    "FRK_Line".Data.BuiltRevision := "FRK_Line".Data.Status.Revision;
    #FRK_DocApply_D011 := TRUE;
END_FUNCTION
FUNCTION "FRK_DocCapture_D012" : Bool
{ S7_Optimized_Access := 'TRUE' }
VERSION : 0.1
VAR_IN_OUT
    Length : DInt;
END_VAR
VAR_TEMP
    Index : Int;
    Stored : Int;
    Position : DInt;
    NativeResult : Int;
    Ok : Bool;
END_VAR
BEGIN
    #FRK_DocCapture_D012 := FALSE;
    "FRK_PersistImages".D012.SchemaVersion := 1; "FRK_PersistImages".D012.Scope := 'PressDemo';
    IF "FRK_ModelRuntime".Rows[1].State = 1 THEN
        #Ok := "FRK_ModelCapture"(RootIndex := 1, Catalog := "FRK_ModelRuntime".Rows[1].Stage, Image := "FRK_PersistImages".D012.Image);
    ELSE
        #Ok := "FRK_ModelCapture"(RootIndex := 1, Catalog := "FRK_ModelStore".Rows[1], Image := "FRK_PersistImages".D012.Image);
    END_IF;
    IF NOT #Ok THEN RETURN; END_IF;
    FOR #Index := 0 TO 2895 DO "FRK_PersistBuffers".D012Data[#Index] := BYTE#0; END_FOR;
    #Position := 24;
    #NativeResult := Serialize(SRC_VARIABLE := "FRK_PersistImages".D012, DEST_ARRAY => "FRK_PersistBuffers".D012Data, POS := #Position);
    IF #NativeResult <> 0 OR #Position < 24 OR #Position > 2896 THEN RETURN; END_IF;
    #Length := #Position - 24;
    #FRK_DocCapture_D012 := TRUE;
END_FUNCTION
FUNCTION "FRK_DocApply_D012" : Bool
{ S7_Optimized_Access := 'TRUE' }
VERSION : 0.1
VAR_TEMP
    Index : Int;
    Stored : Int;
    Position : DInt;
    NativeResult : Int;
    Ok : Bool;
END_VAR
BEGIN
    #FRK_DocApply_D012 := FALSE;
    #Position := 24;
    #NativeResult := Deserialize(SRC_ARRAY := "FRK_PersistBuffers".D012Data, DEST_VARIABLE => "FRK_PersistImages".D012, POS := #Position);
    IF #NativeResult <> 0 OR #Position <> 24 + UDINT_TO_DINT("FRK_PersistConsumers".Rows[12].Result.Length) THEN RETURN; END_IF;
    IF "FRK_PersistImages".D012.SchemaVersion <> 1 OR "FRK_PersistImages".D012.Scope <> 'PressDemo' THEN RETURN; END_IF;
    IF NOT "FRK_ModelApply"(RootIndex := 1, Image := "FRK_PersistImages".D012.Image) THEN RETURN; END_IF;
    #FRK_DocApply_D012 := TRUE;
END_FUNCTION
FUNCTION "FRK_DocReject" : Void
{ S7_Optimized_Access := 'TRUE' }
VERSION : 0.1
VAR_INPUT
    Slot : Int;
END_VAR
VAR_TEMP
    Stored : Int;
END_VAR
BEGIN
    CASE #Slot OF
        1:
            #Stored := "FRK_ConfigFind"(Scope := 'PressDemo', Key := 'degradationPercent', ModelCode := '');
            IF #Stored > 0 THEN "FRK_ConfigStore".Rows[#Stored].Used := FALSE; END_IF;
            #Stored := "FRK_ConfigFind"(Scope := 'PressDemo', Key := 'requireTwoHandStart', ModelCode := '');
            IF #Stored > 0 THEN "FRK_ConfigStore".Rows[#Stored].Used := FALSE; END_IF;
            "FRK_ConfigLoss"(RootIndex := 1, Scope := 'PressDemo');
        2:
            #Stored := "FRK_ConfigFind"(Scope := 'PressDemo', Key := 'idealCycleMs', ModelCode := 'ALUMINUM');
            IF #Stored > 0 THEN "FRK_ConfigStore".Rows[#Stored].Used := FALSE; END_IF;
            #Stored := "FRK_ConfigFind"(Scope := 'PressDemo', Key := 'baselineWorkMs', ModelCode := 'ALUMINUM');
            IF #Stored > 0 THEN "FRK_ConfigStore".Rows[#Stored].Used := FALSE; END_IF;
            #Stored := "FRK_ConfigFind"(Scope := 'PressDemo', Key := 'modeSwitchTimeout', ModelCode := 'ALUMINUM');
            IF #Stored > 0 THEN "FRK_ConfigStore".Rows[#Stored].Used := FALSE; END_IF;
            #Stored := "FRK_ConfigFind"(Scope := 'PressDemo', Key := 'transferSettleTime', ModelCode := 'ALUMINUM');
            IF #Stored > 0 THEN "FRK_ConfigStore".Rows[#Stored].Used := FALSE; END_IF;
            #Stored := "FRK_ConfigFind"(Scope := 'PressDemo', Key := 'pressSettleTime', ModelCode := 'ALUMINUM');
            IF #Stored > 0 THEN "FRK_ConfigStore".Rows[#Stored].Used := FALSE; END_IF;
            "FRK_ConfigLoss"(RootIndex := 1, Scope := 'PressDemo');
        3:
            #Stored := "FRK_ConfigFind"(Scope := 'PressDemo', Key := 'idealCycleMs', ModelCode := 'PLASTIC');
            IF #Stored > 0 THEN "FRK_ConfigStore".Rows[#Stored].Used := FALSE; END_IF;
            #Stored := "FRK_ConfigFind"(Scope := 'PressDemo', Key := 'baselineWorkMs', ModelCode := 'PLASTIC');
            IF #Stored > 0 THEN "FRK_ConfigStore".Rows[#Stored].Used := FALSE; END_IF;
            #Stored := "FRK_ConfigFind"(Scope := 'PressDemo', Key := 'modeSwitchTimeout', ModelCode := 'PLASTIC');
            IF #Stored > 0 THEN "FRK_ConfigStore".Rows[#Stored].Used := FALSE; END_IF;
            #Stored := "FRK_ConfigFind"(Scope := 'PressDemo', Key := 'transferSettleTime', ModelCode := 'PLASTIC');
            IF #Stored > 0 THEN "FRK_ConfigStore".Rows[#Stored].Used := FALSE; END_IF;
            #Stored := "FRK_ConfigFind"(Scope := 'PressDemo', Key := 'pressSettleTime', ModelCode := 'PLASTIC');
            IF #Stored > 0 THEN "FRK_ConfigStore".Rows[#Stored].Used := FALSE; END_IF;
            "FRK_ConfigLoss"(RootIndex := 1, Scope := 'PressDemo');
        4:
            #Stored := "FRK_ConfigFind"(Scope := 'PressDemo', Key := 'idealCycleMs', ModelCode := 'STEEL');
            IF #Stored > 0 THEN "FRK_ConfigStore".Rows[#Stored].Used := FALSE; END_IF;
            #Stored := "FRK_ConfigFind"(Scope := 'PressDemo', Key := 'baselineWorkMs', ModelCode := 'STEEL');
            IF #Stored > 0 THEN "FRK_ConfigStore".Rows[#Stored].Used := FALSE; END_IF;
            #Stored := "FRK_ConfigFind"(Scope := 'PressDemo', Key := 'modeSwitchTimeout', ModelCode := 'STEEL');
            IF #Stored > 0 THEN "FRK_ConfigStore".Rows[#Stored].Used := FALSE; END_IF;
            #Stored := "FRK_ConfigFind"(Scope := 'PressDemo', Key := 'transferSettleTime', ModelCode := 'STEEL');
            IF #Stored > 0 THEN "FRK_ConfigStore".Rows[#Stored].Used := FALSE; END_IF;
            #Stored := "FRK_ConfigFind"(Scope := 'PressDemo', Key := 'pressSettleTime', ModelCode := 'STEEL');
            IF #Stored > 0 THEN "FRK_ConfigStore".Rows[#Stored].Used := FALSE; END_IF;
            "FRK_ConfigLoss"(RootIndex := 1, Scope := 'PressDemo');
        5:
            "FRK_AccessPolicies".Rows[1].Scope := 'PressDemo';
            "FRK_AccessPolicies".Rows[1].SchemaVersion := 0;
            "FRK_AccessPolicies".Rows[1].Initialized := TRUE;
        6:
            "FRK_SetStore".Sets[1, 1].Info.Used := FALSE;
            "FRK_ConfigLoss"(RootIndex := 1, Scope := 'PressDemo');
        7:
            "FRK_SetStore".Sets[1, 2].Info.Used := FALSE;
            "FRK_ConfigLoss"(RootIndex := 1, Scope := 'PressDemo');
        8:
            "FRK_SetStore".Sets[1, 3].Info.Used := FALSE;
            "FRK_ConfigLoss"(RootIndex := 1, Scope := 'PressDemo');
        9:
            "FRK_SetStore".Sets[1, 4].Info.Used := FALSE;
            "FRK_ConfigLoss"(RootIndex := 1, Scope := 'PressDemo');
        10:
            "FRK_LocalUsers".SchemaVersion := 0; "FRK_LocalUsers".Generation := 0; "FRK_LocalUsers".Checksum := DWORD#0;
            "FRK_AccessStorage".UsersCommissioned := TRUE; "FRK_AccessStorage".UsersReady := FALSE; "FRK_AccessStorage".UsersLost := TRUE;
        11:
            "FRK_Line".Data.Dirty := FALSE;
            "FRK_Line".Data.Status.SourceError := 0;
            "FRK_ConfigLoss"(RootIndex := 1, Scope := 'PressDemo');
        12:
            "FRK_ModelStore".Rows[1] := "FRK_ModelRuntime".BlankCatalog;
            "FRK_ModelStore".Rows[1].Scope := 'PressDemo';
            "FRK_ConfigLoss"(RootIndex := 1, Scope := 'PressDemo');
        ELSE RETURN;
    END_CASE;
END_FUNCTION
FUNCTION "FRK_DocCapture" : Void
{ S7_Optimized_Access := 'TRUE' }
VERSION : 0.1
VAR_INPUT
    Slot : Int;
END_VAR
VAR_IN_OUT
    Ok : Bool;
    Length : DInt;
END_VAR
BEGIN
    #Ok := FALSE; #Length := 0;
    CASE #Slot OF
        1: #Ok := "FRK_DocCapture_D001"(Length := #Length);
        2: #Ok := "FRK_DocCapture_D002"(Length := #Length);
        3: #Ok := "FRK_DocCapture_D003"(Length := #Length);
        4: #Ok := "FRK_DocCapture_D004"(Length := #Length);
        5: #Ok := "FRK_DocCapture_D005"(Length := #Length);
        6: #Ok := "FRK_DocCapture_D006"(Length := #Length);
        7: #Ok := "FRK_DocCapture_D007"(Length := #Length);
        8: #Ok := "FRK_DocCapture_D008"(Length := #Length);
        9: #Ok := "FRK_DocCapture_D009"(Length := #Length);
        10: #Ok := "FRK_DocCapture_D010"(Length := #Length);
        11: #Ok := "FRK_DocCapture_D011"(Length := #Length);
        12: #Ok := "FRK_DocCapture_D012"(Length := #Length);
        ELSE RETURN;
    END_CASE;
END_FUNCTION
FUNCTION "FRK_DocApply" : Bool
{ S7_Optimized_Access := 'TRUE' }
VERSION : 0.1
VAR_INPUT
    Slot : Int;
END_VAR
BEGIN
    #FRK_DocApply := FALSE;
    CASE #Slot OF
        1: #FRK_DocApply := "FRK_DocApply_D001"();
        2: #FRK_DocApply := "FRK_DocApply_D002"();
        3: #FRK_DocApply := "FRK_DocApply_D003"();
        4: #FRK_DocApply := "FRK_DocApply_D004"();
        5: #FRK_DocApply := "FRK_DocApply_D005"();
        6: #FRK_DocApply := "FRK_DocApply_D006"();
        7: #FRK_DocApply := "FRK_DocApply_D007"();
        8: #FRK_DocApply := "FRK_DocApply_D008"();
        9: #FRK_DocApply := "FRK_DocApply_D009"();
        10: #FRK_DocApply := "FRK_DocApply_D010"();
        11: #FRK_DocApply := "FRK_DocApply_D011"();
        12: #FRK_DocApply := "FRK_DocApply_D012"();
        ELSE RETURN;
    END_CASE;
END_FUNCTION
FUNCTION "FRK_DocBoot" : Void
{ S7_Optimized_Access := 'TRUE' }
VERSION : 0.1
VAR_INPUT
    Startup : Bool;
END_VAR
VAR_IN_OUT
    Ready : Bool;
END_VAR
VAR_TEMP
    Slot : Int;
    Done : Bool;
    Ok : Bool;
END_VAR
BEGIN
    IF #Startup THEN
        "FRK_PersistConsumers".Ready := FALSE;
        FOR #Slot := 1 TO 12 DO
            "FRK_PersistConsumers".Rows[#Slot].State := 0; "FRK_PersistConsumers".Rows[#Slot].Ticket := 0;
            "FRK_PersistConsumers".Rows[#Slot].Dirty := FALSE; "FRK_PersistConsumers".Rows[#Slot].Failed := FALSE;
            "FRK_PersistConsumers".Rows[#Slot].Rejected := FALSE; "FRK_PersistConsumers".Rows[#Slot].Acknowledged := FALSE;
            "FRK_PersistConsumers".Rows[#Slot].RetrySince := "FRK_Clock".NowMs;
            "FRK_PersistConsumers".Rows[#Slot].PendingSince := LDT#1970-01-01-00:00:00;
            "FRK_PersistConsumers".Rows[#Slot].NextSince := LDT#1970-01-01-00:00:00;
        END_FOR;
    END_IF;
    #Ready := TRUE;
    "FRK_PersistStatus".Failed := FALSE;
    FOR #Slot := 1 TO 12 DO
        IF "FRK_PersistConsumers".Rows[#Slot].State = 0 THEN
            IF NOT "FRK_PersistConsumers".Rows[#Slot].Failed OR "FRK_Elapsed"(NewMs := "FRK_Clock".NowMs, OldMs := "FRK_PersistConsumers".Rows[#Slot].RetrySince) >= 1000 THEN
                "FRK_PersistConsumers".Rows[#Slot].Ticket := "FRK_PersistStart"(Slot := #Slot, WriteDocument := FALSE, Length := 0);
                IF "FRK_PersistConsumers".Rows[#Slot].Ticket <> 0 THEN "FRK_PersistConsumers".Rows[#Slot].State := 1; END_IF;
            END_IF;
        ELSIF "FRK_PersistConsumers".Rows[#Slot].State = 1 THEN
            #Done := "FRK_PersistPoll"(Ticket := "FRK_PersistConsumers".Rows[#Slot].Ticket, Result := "FRK_PersistConsumers".Rows[#Slot].Result);
            IF #Done THEN
                "FRK_PersistConsumers".Rows[#Slot].Ticket := 0;
                IF NOT "FRK_PersistConsumers".Rows[#Slot].Result.Ok THEN
                    "FRK_PersistConsumers".Rows[#Slot].Failed := TRUE; "FRK_PersistConsumers".Rows[#Slot].State := 0;
                    "FRK_PersistConsumers".Rows[#Slot].RetrySince := "FRK_Clock".NowMs;
                ELSE
                    "FRK_PersistConsumers".Rows[#Slot].Failed := FALSE;
                    #Ok := NOT "FRK_PersistConsumers".Rows[#Slot].Result.Lost;
                    "FRK_PersistConsumers".Rows[#Slot].Virgin := #Ok AND NOT "FRK_PersistConsumers".Rows[#Slot].Result.Found;
                    IF #Ok AND "FRK_PersistConsumers".Rows[#Slot].Result.Found THEN #Ok := "FRK_DocApply"(Slot := #Slot); END_IF;
                    IF NOT #Ok THEN
                        "FRK_DocReject"(Slot := #Slot);
                        "FRK_PersistConsumers".Rows[#Slot].Rejected := TRUE;
                    ELSIF "FRK_PersistConsumers".Rows[#Slot].Virgin THEN "FRK_PersistDirty"(Slot := #Slot); END_IF;
                    "FRK_PersistConsumers".Rows[#Slot].State := 2;
                END_IF;
            END_IF;
        END_IF;
        IF "FRK_PersistConsumers".Rows[#Slot].State <> 2 THEN #Ready := FALSE; END_IF;
        "FRK_PersistStatus".Failed := "FRK_PersistStatus".Failed OR "FRK_PersistConsumers".Rows[#Slot].Failed;
    END_FOR;
    "FRK_PersistStatus".Restoring := NOT #Ready;
    "FRK_PersistStatus".NativeStatus := INT_TO_WORD("FRK_PersistRuntime".NativeResult);
    "FRK_PersistConsumers".Ready := #Ready;
END_FUNCTION
FUNCTION "FRK_DocCyclic" : Void
{ S7_Optimized_Access := 'TRUE' }
VERSION : 0.1
VAR_TEMP
    Slot : Int;
    Done : Bool;
    Ok : Bool;
    Length : DInt;
END_VAR
BEGIN
    IF NOT "FRK_PersistConsumers".Ready THEN RETURN; END_IF;
    FOR #Slot := 1 TO 12 DO
        IF "FRK_PersistConsumers".Rows[#Slot].Ticket <> 0 THEN
            #Done := "FRK_PersistPoll"(Ticket := "FRK_PersistConsumers".Rows[#Slot].Ticket, Result := "FRK_PersistConsumers".Rows[#Slot].Result);
            IF #Done THEN
                "FRK_PersistConsumers".Rows[#Slot].Ticket := 0;
                "FRK_PersistConsumers".Rows[#Slot].Failed := NOT "FRK_PersistConsumers".Rows[#Slot].Result.Ok;
                "FRK_PersistConsumers".Rows[#Slot].RetrySince := "FRK_Clock".NowMs;
                IF "FRK_PersistConsumers".Rows[#Slot].Failed THEN "FRK_PersistConsumers".Rows[#Slot].Dirty := TRUE;
                ELSIF "FRK_PersistConsumers".Rows[#Slot].Dirty THEN "FRK_PersistConsumers".Rows[#Slot].PendingSince := "FRK_PersistConsumers".Rows[#Slot].NextSince;
                ELSE "FRK_PersistConsumers".Rows[#Slot].PendingSince := LDT#1970-01-01-00:00:00; END_IF;
            END_IF;
        ELSIF "FRK_PersistConsumers".Rows[#Slot].Dirty AND (NOT "FRK_PersistConsumers".Rows[#Slot].Rejected OR "FRK_PersistConsumers".Rows[#Slot].Acknowledged) THEN
            IF NOT "FRK_PersistConsumers".Rows[#Slot].Failed OR "FRK_Elapsed"(NewMs := "FRK_Clock".NowMs, OldMs := "FRK_PersistConsumers".Rows[#Slot].RetrySince) >= 1000 THEN
                "FRK_DocCapture"(Slot := #Slot, Ok := #Ok, Length := #Length);
                IF #Ok THEN
                    "FRK_PersistConsumers".Rows[#Slot].Ticket := "FRK_PersistStart"(Slot := #Slot, WriteDocument := TRUE, Length := #Length);
                    IF "FRK_PersistConsumers".Rows[#Slot].Ticket <> 0 THEN "FRK_PersistConsumers".Rows[#Slot].Dirty := FALSE; END_IF;
                ELSE "FRK_PersistConsumers".Rows[#Slot].Failed := TRUE; "FRK_PersistConsumers".Rows[#Slot].RetrySince := "FRK_Clock".NowMs; END_IF;
            END_IF;
        END_IF;
    END_FOR;
END_FUNCTION
